FUNCTION_BLOCK FaseAtivaNereda (* Numero da fase ativa e da fase abortada (pela ordem das entradas) e indicacao de abortado *)
  (* Standard: 61499-2 *)
  (* Version 1.1, 05/11/2026, Hidryco, Hidryco, 1.1: fase ativa = Starting OU Run OU Stopping OU Aborting (entradas PartindoN, ParandoN, AbortandoN). 1.0: FaseAtiva = numero da 1a entrada RunN em TRUE (0 = nenhuma); FaseAbortada = numero da 1a AbortadaN em TRUE (0 = nenhuma); Abortado = alguma AbortadaN. CNF so quando muda (e na 1a execucao). Eventos de saida no ECAction. *)
  PACKAGE SE.Nereda;
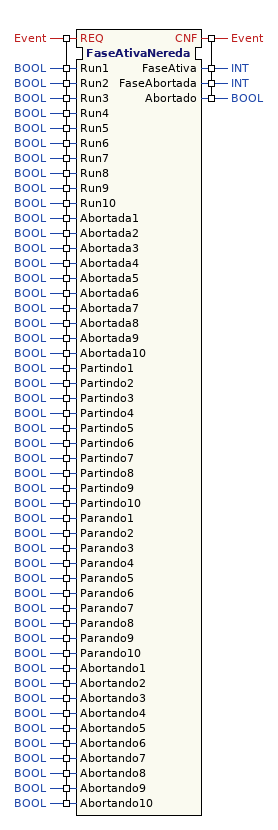
  EVENT_INPUT
    REQ WITH Run1, Run2, Run3, Run4, Run5, Run6, Run7, Run8, Run9, Run10, Abortada1, Abortada2, Abortada3, Abortada4, Abortada5, Abortada6, Abortada7, Abortada8, Abortada9, Abortada10, Partindo1, Partindo2, Partindo3, Partindo4, Partindo5, Partindo6, Partindo7, Partindo8, Partindo9, Partindo10, Parando1, Parando2, Parando3, Parando4, Parando5, Parando6, Parando7, Parando8, Parando9, Parando10, Abortando1, Abortando2, Abortando3, Abortando4, Abortando5, Abortando6, Abortando7, Abortando8, Abortando9, Abortando10; (* Estado das fases mudou *)
  END_EVENT
  EVENT_OUTPUT
    CNF WITH FaseAtiva, FaseAbortada, Abortado; (* Fase ativa ou abortada mudou *)
  END_EVENT
  VAR_INPUT
    Run1 : BOOL; (* Fase 1 rodando *)
    Run2 : BOOL; (* Fase 2 rodando *)
    Run3 : BOOL; (* Fase 3 rodando *)
    Run4 : BOOL; (* Fase 4 rodando *)
    Run5 : BOOL; (* Fase 5 rodando *)
    Run6 : BOOL; (* Fase 6 rodando *)
    Run7 : BOOL; (* Fase 7 rodando *)
    Run8 : BOOL; (* Fase 8 rodando *)
    Run9 : BOOL; (* Fase 9 rodando *)
    Run10 : BOOL; (* Fase 10 rodando *)
    Abortada1 : BOOL; (* Fase 1 abortada *)
    Abortada2 : BOOL; (* Fase 2 abortada *)
    Abortada3 : BOOL; (* Fase 3 abortada *)
    Abortada4 : BOOL; (* Fase 4 abortada *)
    Abortada5 : BOOL; (* Fase 5 abortada *)
    Abortada6 : BOOL; (* Fase 6 abortada *)
    Abortada7 : BOOL; (* Fase 7 abortada *)
    Abortada8 : BOOL; (* Fase 8 abortada *)
    Abortada9 : BOOL; (* Fase 9 abortada *)
    Abortada10 : BOOL; (* Fase 10 abortada *)
    Partindo1 : BOOL; (* Fase 1 em Starting *)
    Partindo2 : BOOL; (* Fase 2 em Starting *)
    Partindo3 : BOOL; (* Fase 3 em Starting *)
    Partindo4 : BOOL; (* Fase 4 em Starting *)
    Partindo5 : BOOL; (* Fase 5 em Starting *)
    Partindo6 : BOOL; (* Fase 6 em Starting *)
    Partindo7 : BOOL; (* Fase 7 em Starting *)
    Partindo8 : BOOL; (* Fase 8 em Starting *)
    Partindo9 : BOOL; (* Fase 9 em Starting *)
    Partindo10 : BOOL; (* Fase 10 em Starting *)
    Parando1 : BOOL; (* Fase 1 em Stopping *)
    Parando2 : BOOL; (* Fase 2 em Stopping *)
    Parando3 : BOOL; (* Fase 3 em Stopping *)
    Parando4 : BOOL; (* Fase 4 em Stopping *)
    Parando5 : BOOL; (* Fase 5 em Stopping *)
    Parando6 : BOOL; (* Fase 6 em Stopping *)
    Parando7 : BOOL; (* Fase 7 em Stopping *)
    Parando8 : BOOL; (* Fase 8 em Stopping *)
    Parando9 : BOOL; (* Fase 9 em Stopping *)
    Parando10 : BOOL; (* Fase 10 em Stopping *)
    Abortando1 : BOOL; (* Fase 1 em Aborting *)
    Abortando2 : BOOL; (* Fase 2 em Aborting *)
    Abortando3 : BOOL; (* Fase 3 em Aborting *)
    Abortando4 : BOOL; (* Fase 4 em Aborting *)
    Abortando5 : BOOL; (* Fase 5 em Aborting *)
    Abortando6 : BOOL; (* Fase 6 em Aborting *)
    Abortando7 : BOOL; (* Fase 7 em Aborting *)
    Abortando8 : BOOL; (* Fase 8 em Aborting *)
    Abortando9 : BOOL; (* Fase 9 em Aborting *)
    Abortando10 : BOOL; (* Fase 10 em Aborting *)
  END_VAR
  VAR_OUTPUT
    FaseAtiva : INT; (* 0 = nenhuma; N = fase da entrada RunN *)
    FaseAbortada : INT; (* 0 = nenhuma; N = fase da entrada AbortadaN *)
    Abortado : BOOL; (* TRUE = alguma fase abortada *)
  END_VAR
  VAR
    primeira : BOOL := TRUE; (* Forca o CNF na 1a execucao *)
    oldFaseAtiva : INT;
    oldFaseAbortada : INT;
    oldAbortado : BOOL;
  END_VAR
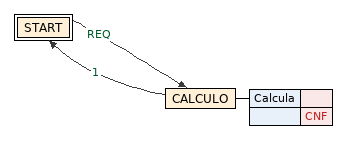
  EC_STATES
    START; (* Estado inicial *)
    CALCULO : Calcula, -> CNF; (* Calcula; CNF so quando muda *)
  END_STATES
  EC_TRANSITIONS
    START TO CALCULO := REQ;
    CALCULO TO START := 1;
  END_TRANSITIONS
  ALGORITHM Calcula IN ST: (* Numero da fase ativa e da abortada *)
CNF := FALSE;
IF (Run1 OR Partindo1 OR Parando1 OR Abortando1) THEN
    FaseAtiva := 1;
ELSIF (Run2 OR Partindo2 OR Parando2 OR Abortando2) THEN
    FaseAtiva := 2;
ELSIF (Run3 OR Partindo3 OR Parando3 OR Abortando3) THEN
    FaseAtiva := 3;
ELSIF (Run4 OR Partindo4 OR Parando4 OR Abortando4) THEN
    FaseAtiva := 4;
ELSIF (Run5 OR Partindo5 OR Parando5 OR Abortando5) THEN
    FaseAtiva := 5;
ELSIF (Run6 OR Partindo6 OR Parando6 OR Abortando6) THEN
    FaseAtiva := 6;
ELSIF (Run7 OR Partindo7 OR Parando7 OR Abortando7) THEN
    FaseAtiva := 7;
ELSIF (Run8 OR Partindo8 OR Parando8 OR Abortando8) THEN
    FaseAtiva := 8;
ELSIF (Run9 OR Partindo9 OR Parando9 OR Abortando9) THEN
    FaseAtiva := 9;
ELSIF (Run10 OR Partindo10 OR Parando10 OR Abortando10) THEN
    FaseAtiva := 10;
ELSE
    FaseAtiva := 0;
END_IF;
IF Abortada1 THEN
    FaseAbortada := 1;
ELSIF Abortada2 THEN
    FaseAbortada := 2;
ELSIF Abortada3 THEN
    FaseAbortada := 3;
ELSIF Abortada4 THEN
    FaseAbortada := 4;
ELSIF Abortada5 THEN
    FaseAbortada := 5;
ELSIF Abortada6 THEN
    FaseAbortada := 6;
ELSIF Abortada7 THEN
    FaseAbortada := 7;
ELSIF Abortada8 THEN
    FaseAbortada := 8;
ELSIF Abortada9 THEN
    FaseAbortada := 9;
ELSIF Abortada10 THEN
    FaseAbortada := 10;
ELSE
    FaseAbortada := 0;
END_IF;
Abortado := FaseAbortada <> 0;
CNF := primeira OR (FaseAtiva <> oldFaseAtiva) OR (FaseAbortada <> oldFaseAbortada) OR (Abortado <> oldAbortado);
primeira := FALSE;
oldFaseAtiva := FaseAtiva;
oldFaseAbortada := FaseAbortada;
oldAbortado := Abortado;
  END_ALGORITHM
END_FUNCTION_BLOCK
